(*
SPDX-FileCopyrightText: © 2026 Oleksandr Tiutyk <trofimich@gmail.com>
SPDX-License-Identifier: MIT
License: https://opensource.org/license/mit
*)

(*!
<summary>Stores an owned text snapshot waiting for a logging backend.</summary>
<description>
Internal QueuedLogger storage. Text, category and optional number are copied by value. Contains no borrowed
references to caller data or exceptions.
</description>
*)
TYPE QUEUED_LOG_MESSAGE :
STRUCT
	Message : TOF_Core.ERROR_MESSAGE;
	Category : TOF_Core.LOG_CATEGORY;
	HasMessageNumber : BOOL;
	MessageNumber : ULINT;
END_STRUCT
END_TYPE

(* stored: Version 1.1.0.1
   DUT QUEUED_LOG_MESSAGE: Id {351add95-024d-43b6-b667-88459d6b5588} *)
